//---------------------------------------------------------------------------------------------------------------
//
//  HAUD 2026.11.23
//
//
//---------------------------------------------------------------------------------------------------------------
//  fb_Instance
//---------------------------------------------------------------------------------------------------------------
//---------------------------------------------------------------------------------------------------------------
//  - base class for a process instance to work with fb_ProcessCollector
//  - extend this class to build top level transport logic
//    - example extension: fb_DistributorByTicket (1 to many)
//
//  What is it that I truly desire? 
//  --> to reduce the amount of handshakes that are required for a range of XtsStation
//  --> keep the granularity of a single station also for a range of stations
//  --> reuse existing interfaces
//
//  What an Instance is for:
//  - customized administrative transport related work
//    - reading of process tickets
//    - checking of queues
//    - handshaking ranges of stations
//      - automate handshake sequences with the collectors
//    - letting the stations write station tickets
//    - writing of process tickets
//
//  How an Instance is supposed to work:
//  - An Instance is of the same nature as a fb_StationProcess.Cycle / fb_ProcessCollector.Cycle
//    
//    --> you should build a Cycle() method
//    --> the default state after self init at PowerOn shall be a disabled state
//      --> a station behaviour follows the following concept:
//        - switch on --> station moves to enabled state
//        - enabled : switch to detection
//          - detection : detect what is given to you (e.g. QueueCount or LinkedList ticket)
//          - detected work leads to station asking for permission
//        - permitted : execute whatever is mandatory for starting the process (move to position etc)
//        - start / done
//          --> you decide how to handshake
//        - ready to send out : prepare your destination data here!
//        - send out : handshake sequence for safely permitting motion of a mover and transport of information
//
//    - It is up to you to decide how many handshakes with the CollectorInterface to automate in an instance
//      - example, a default distributor may require handshakes for every mover, 
//                 a mask driven distributor distributes until it has worked through the mask autonomously
//
//    - Read the existing extensions:
//      - you will find a 2-step progression for state changes
//      - they use the enumerations E_INSTANCE_CMD / E_INSTANCE_STATE
//        - in combination with E_PROGRESS
//        - there will be flowcharts for the existing extensions.
//
//---------------------------------------------------------------------------------------------------------------
//  - there are already 3 primitives available
//    - [1 to 1] DistributorByQueue
//      - a single station for 
//        - fly-by and change dynamics
//        - simple one stop
//
//    - [1 to m] DistributorByTicket
//      - a single station with ticket inbox check for
//        - sending a mover to a range of stations in accordance to the bitmask it received
//
//    - [m to 1] ProcessByTicket
//      - a range of stations handling a stationary process with ticket inbox
//      - single and nested stops
//      - sends movers to a single target (distributor)
//---------------------------------------------------------------------------------------------------------------
//
//---------------------------------------------------------------------------------------------------------------
//  - ProcessId : _nProcess --> whoami, this is me
//---------------------------------------------------------------------------------------------------------------
//
//  - who is required for my work on the outside?
//  - fb_ProcessCollector[_nProcess].Cycle() is called in MAIN_APP(PRG)
//    - provides interface
//    - handles range of XtsStations
//    - range must be closed and in consecutive order
//
//    - combines states into bitmasks, one bit per XtsStation
//    - controls forwarding of commands to range of XtsStations 
//      (see fb_ProcessCollector.Cycle())
//
//---------------------------------------------------------------------------------------------------------------
//  - CollectorInterface 
//---------------------------------------------------------------------------------------------------------------
//    - reference to all _ItfProcessCollector(I_ProcessCollector)[]
//    - _ItfProcessCollector[nProcess] carries ctrl/state information
//
//    - Control / State of the CollectorInterface
//      - local _stCollectorCtrl / _stCollectorState datafields are linked (REF=) to CollectorInterface.ProcessCtrl / .ProcessState
//        - since this connection shall be done automatically I put it in Check() method
//          --> see Check()
// 
//      - local datafield for control and state provided
//        - since CollectorInterface.ProcessCtrl and CollectorInterface.ProcessState are reference pointers
//          --> the real datafield has to come from somewhere, 
//              in this case the local datafields _stCollectorCtrl/_stCollectorState
//
//      - _stCollectorCtrl(ST_PROCESS_CTRL)
//        --> commands to the connected CollectorInterface;
//
//        Cmd               : E_PROCESS_CTRL; // command enum for collector
//        ProcessTarget     : UINT;           // target of my process
//        ActivateStation   : T_PROCESS;      // is checked for every job
//                                            // every bit is an XtsStation
//
//        NestMask          : BYTE;           // one mask for all XtsStations
//        - every bit is a PosStop within an XtsStation
//
//      - _stCollectorState(ST_PROCESS_STATE)
//        --> status information from the connected CollectorInterface
//        --> check for plausible StationLast / StationFirst range of XtsStations
//
//        State             : E_PROCESS_STATE;  // state enum from collector
//        Result            : E_PROGRESS;       // substate from collector, E_PROGRESS.PROGRESS_BUSY signals the collector state is ready for interaction
//                                              // fb_DistributorByTicket may give you an idea of the use of a substate 
//        Check             : E_PROCESS_CHECK;  // plausibility check of StationLast and StationFirst (the result of Check() --> _eCheck) 
//---------------------------------------------------------------------------------------------------------------
//  - InstanceCtrl(_stInstanceCtrl) 
//---------------------------------------------------------------------------------------------------------------
//  - incoming handshakes from higher up
//    - remember, 
//      this shall be a helper so you can do administrative stuff here 
//      so your actual process logic (picking, dispensing, syncing, gearing) may live elsewhere
// 
//---------------------------------------------------------------------------------------------------------------
//  - InstanceState(_stInstanceState)
//---------------------------------------------------------------------------------------------------------------
//  - reporting to higher up
//
//
//---------------------------------------------------------------------------------------------------------------
//---------------------------------------------------------------------------------------------------------------
//  - basic check and var names, so you can build your procedures with it
//
//  - processes may be connected via linked list, you decide.
//    - linked list for processes is intended to work as job buffer
//    - linked list provides information via ST_PROCESS_DATA, 
//      add what you have to in there
//    - linked list to all process instances provided
//
//  - inherit this base class for your application, call Check() every cycle at the top before you do anything
//       IF NOT Check() THEN 
//         RETURN; 
//       END_IF
//
//---------------------------------------------------------------------------------------------------------------//
// This SOFTWARE is provided as an Example by THE PROVIDER "as is" and "with all faults." THE PROVIDER makes no  //
// representations or warranties of any kind concerning the safety, suitability, lack of viruses, inaccuracies,  //
// typographical errors, or other harmful components of this SOFTWARE. There are inherent dangers in the use of  //
// any software, and you are solely responsible for determining whether this SOFTWARE is compatible with your    //
// equipment and other software installed on your equipment. You are also solely responsible for the protection  //
// of your equipment and backup of your data, and THE PROVIDER will not be liable for any damages you may suffer //
// in connection with using, modifying, or distributing this SOFTWARE.                                           //
//---------------------------------------------------------------------------------------------------------------//
FUNCTION_BLOCK ABSTRACT fb_Instance
VAR
  // process index
  _nProcess               : E_INSTANCE;           // whoami

  _stInstanceCtrl         : REFERENCE TO ARRAY[1..MAX_PROCESS] OF ST_INSTANCE_CTRL;
  _stInstanceState        : REFERENCE TO ARRAY[1..MAX_PROCESS] OF ST_INSTANCE_STATE;

  _eCmd,
  _eCmdOld                : E_INSTANCE_CMD;       // commands for local state machine
  _eStateInstance         : E_INSTANCE_STATE;     // local state machine for infeed procedure

  _eResult                : E_PROGRESS;           // result for methods
  _eStateProgress         : E_PROGRESS;           // substate for local state machine

  _eInit                  : E_PROGRESS;           // startup
  _eCheck                 : E_INSTANCE_CHECK;     // pointer checks

  // local ctrl / state datafields for you to use, connected by reference to _ItfProcessCollector[_nProcess]
  _stCollectorCtrl        : ST_PROCESS_CTRL;      // control to write, connected by reference to _ItfProcessCollector
  _stCollectorState       : ST_PROCESS_STATE;     // state   to read,  connected by reference to _ItfProcessCollector

  _ItfProcessCollector    : ARRAY[1..MAX_PROCESS] OF I_ProcessCollector;    // information and configuration of the connected ProcessCollector for given range of XtsStations

  _ItfProcessList         : ARRAY[1..MAX_PROCESS] OF I_Process_LinkedList;  // access to all linked lists for writing tickets
  _stListResult           : ST_PROCESS_LIST_RESULT;
  _stProcessData          : ST_PROCESS_DATA;

  {attribute 'displaymode':='bin'}
  _wTargetMask            : ARRAY[1..SIZEOF(T_PROCESS)*8] OF BYTE; // bits for PosStop[] to use in XtsStation of target process

  // position window within which a mover must be for the instance to react
  // value in abs modulo axis value
  //  - crossing the modulo turn is evaluated --> (Start > End) case is valid as window
  _rCheckPositionStart    : LREAL;
  _rCheckPositionEnd      : LREAL;

  _stMsg                  : ST_Message;
  _MessageLevel           : E_MessageType := E_MessageType.eMessageInfo;
END_VAR

METHOD Check : BOOL // call this method in the extending/inheriting class
//-----------------------------------------------------------------------------
//-----------------------------------------------------------------------------
// plausibility checks
//-----------------------------------------------------------------------------
IF NOT (_nProcess > 0)
THEN
  _eCheck                 := E_INSTANCE_CHECK.PROCESS_ID_ZERO;
  RETURN;
END_IF

IF NOT (_nProcess < E_INSTANCE.INSTANCE_MAX)
THEN
  _eCheck                 := E_INSTANCE_CHECK.PROCESS_ID_MAX;
  RETURN;
END_IF
//-----------------------------------------------------------------------------
//-----------------------------------------------------------------------------
// pointer checks
//-----------------------------------------------------------------------------
IF NOT __ISVALIDREF(_stInstanceCtrl)
THEN
  _eCheck                 := E_INSTANCE_CHECK.INVALID_INSTANCE_CONTROL_REFERENCE;
  RETURN;
END_IF

IF NOT __ISVALIDREF(_stInstanceState)
THEN
  _eCheck                 := E_INSTANCE_CHECK.INVALID_INSTANCE_STATE_REFERENCE;
  RETURN;
END_IF

IF NOT (_ItfProcessCollector[_nProcess] <> 0) 
THEN
  _eCheck                 := E_INSTANCE_CHECK.POINTER_COLLECTOR_ITF_INVALID;
  RETURN;
END_IF

IF NOT (_ItfProcessCollector[_nProcess].ProcessId > 0)
THEN
  _eCheck                 := E_INSTANCE_CHECK.PROCESS_ID_ZERO;
  RETURN;
END_IF

IF NOT (_ItfProcessCollector[_nProcess].ProcessId < E_INSTANCE.INSTANCE_MAX)
THEN
  _eCheck                 := E_INSTANCE_CHECK.PROCESS_ID_MAX;
  RETURN;
END_IF

IF NOT (_nProcess = _ItfProcessCollector[_nProcess].ProcessId)
THEN
  _eCheck                 := E_INSTANCE_CHECK.PROCESS_ID_NOTEQUAL_COLLECTOR_ID;
  RETURN;
END_IF

IF NOT (_ItfProcessList[_nProcess] <> 0)
THEN
  _eCheck                 := E_INSTANCE_CHECK.PROCESS_LIST_ITF_INDEX_INVALID;
  RETURN;
END_IF
//-----------------------------------------------------------------------------
//-----------------------------------------------------------------------------
// connect datafields to interface of ProcessCollector
//-----------------------------------------------------------------------------
_ItfProcessCollector[_nProcess].ProcessCtrl   REF= _stCollectorCtrl;
_ItfProcessCollector[_nProcess].ProcessState  REF= _stCollectorState;

//-----------------------------------------------------------------------------
//-----------------------------------------------------------------------------
// set message device
//-----------------------------------------------------------------------------
_stMsg.eDevice            := e_Device.Process + TO_UINT(_nProcess);
//-----------------------------------------------------------------------------
//-----------------------------------------------------------------------------
_eCheck                   := E_INSTANCE_CHECK.CHECK_DONE;
Check                     := TRUE;
END_METHOD

PROPERTY CheckPositionEnd : lreal // end of the position window to execute logic (should be higher than the WaitPos this instance is working on)
GET
CheckPositionEnd := _rCheckPositionEnd;
END_GET
SET
_rCheckPositionEnd := CheckPositionEnd;
END_SET
END_PROPERTY

PROPERTY CheckPositionStart : lreal // start of the position window to execute instance logic
GET
CheckPositionStart := _rCheckPositionStart;
END_GET
SET
_rCheckPositionStart := CheckPositionStart;
END_SET
END_PROPERTY

METHOD CmdLog

IF (_MessageLevel > E_MessageType.eMessageError)
THEN
  _stMsg.eSubdevice       := e_Subdevice.Instance_Command;
  _stMsg.iErrorNumber     := _nProcess;
  _stMsg.sText            := concat('E_INSTANCE_CMD', '.');
  _stMsg.sText            := concat(_stMsg.sText, TO_STRING(_eCmd));
  f_MessageSet(_stMsg);
END_IF
END_METHOD

PROPERTY CollectorInterface : array[1..MAX_PROCESS] of I_ProcessCollector
SET
_ItfProcessCollector := CollectorInterface;
END_SET
END_PROPERTY

PROPERTY InstanceCtrl : REFERENCE TO ARRAY[1..MAX_PROCESS] OF ST_INSTANCE_CTRL
SET
_stInstanceCtrl ref= InstanceCtrl;
END_SET
END_PROPERTY

PROPERTY InstanceState : REFERENCE TO ARRAY[1..MAX_PROCESS] OF ST_INSTANCE_STATE
SET
_stInstanceState ref= InstanceState;
END_SET
END_PROPERTY

PROPERTY MessageLevel : e_MessageType
GET
MessageLevel := _MessageLevel;
END_GET
SET
_MessageLevel := MessageLevel;

IF NOT (_eInit  = E_PROGRESS.PROGRESS_DONE) OR
   NOT (_eCheck = E_INSTANCE_CHECK.CHECK_DONE)
THEN
  RETURN;
ELSE
  _ItfProcessCollector[_nProcess].MessageLevel := _MessageLevel;
END_IF
END_SET
END_PROPERTY

PROPERTY ProcessId : E_INSTANCE
GET
ProcessId := _nProcess;
END_GET
SET
_nProcess := ProcessId;
END_SET
END_PROPERTY

PROPERTY ProcessLinkedLists : ARRAY[1..max_process] OF I_Process_LinkedList
SET
_ItfProcessList := ProcessLinkedLists;
END_SET
END_PROPERTY

END_FUNCTION_BLOCK

(* stored: Version 1.1.0.1
   POU fb_Instance: Id {aa404a3e-1847-48a0-90da-b76021166e7c}, SpecialFunc None
   Folder properties: Id {3fc25e2e-f78a-4e4b-8f93-14def1aa86a2}
   Method Check: Id {9cd29f0b-abaf-4789-854c-ec925ea6b0ca}
   Property CheckPositionEnd: Id {611133ef-1aa7-4cac-8c52-cbfc3d44858b}
   Get Get: Id {220e427a-8106-496d-8e02-efe34fe069d3}
   Set Set: Id {3c54014d-4c7a-4e01-845f-ae2fc227ec95}
   Property CheckPositionStart: Id {74147dd9-e508-4775-99ef-aeb3905c9fab}
   Get Get: Id {02431a8b-a3c4-49ec-816f-3fbbb6eb28a7}
   Set Set: Id {49a13307-7d3e-4cb3-a294-b3105053b320}
   Method CmdLog: Id {59b1c5ef-8900-4988-bf5d-ece023138df6}
   Property CollectorInterface: Id {1778065e-71fc-4b61-95e9-f0ce7344fd52}
   Set Set: Id {efa86bb5-063c-45e0-824e-e0c7dd62a865}
   Property InstanceCtrl: Id {981757e0-8e40-45aa-8057-0491d6ad023f}
   Set Set: Id {c8e80f92-c362-4f41-b0f9-db9dbea0e4aa}
   Property InstanceState: Id {c8bdcdf1-4ecd-4637-8eac-c66b80a81d6a}
   Set Set: Id {03b5b73e-3a6b-4866-9a71-452e2580c4e5}
   Property MessageLevel: Id {14a41416-0811-40c7-bca5-c73484c900e8}
   Get Get: Id {55960fd5-ef50-4cb1-ac26-92fb20141955}
   Set Set: Id {919b1481-002a-4dbe-8ca4-b1c293d8d704}
   Property ProcessId: Id {0e2c48f6-df86-4fbb-8e57-b52b71d7cbbe}
   Get Get: Id {f8401d20-eb74-43d4-9fe4-3c8cf8a9917e}
   Set Set: Id {a4eb999b-e525-42f5-b031-b3d17e5e8ef9}
   Property ProcessLinkedLists: Id {2f89974a-bbab-4971-8579-59c8d4c1391a}
   Set Set: Id {f0e2969e-ffb1-4ccd-ace6-2a5cd31e132b} *)
